(*!
<summary>Provides floating-point and raw-bit views of the same 32-bit storage.</summary>
<description>
Value and Raw overlap. Reading the other member reinterprets bits; it does not perform numeric conversion.
</description>
*)
TYPE REAL_UNION :
UNION
    Value : REAL;
    Raw : UDINT;
END_UNION
END_TYPE

(* stored: Version 1.1.0.1
   DUT REAL_UNION: Id {45a8f752-e352-42e7-996a-402c3a7b3513} *)
